// TIA Portal V20 export
// export: Created 2026-10-12T15:46:51.9760666Z, ExportSetting WithDefaults, DisplayName Totally Integrated Automation Portal, DisplayVersion V20, DisplayName TIA Portal Openness, DisplayVersion V20, DisplayName TIA Portal Teamcenter Gateway, DisplayVersion V20, DisplayName TIA Portal Version Control Interface, DisplayVersion V20, DisplayName SINAMICS Startdrive Advanced, DisplayVersion V20 SP1 Update 2, DisplayName SINAMICS Startdrive G110M, G120, G120C, G120D, G120P, G115D, DisplayVersion V20 SP1 Update 2, DisplayName SINAMICS Startdrive G130, G150, S120, S150, SINAMICS MV, G220, S200, S210, DisplayVersion V20 SP1 Update 2, DisplayName STEP 7 Professional, DisplayVersion V20, DisplayName STEP 7 Safety, DisplayVersion V20, DisplayName WinCC Basic/Comfort/Advanced, DisplayVersion V20, DisplayName WinCC Professional, DisplayVersion V20, DisplayName WinCC Unified, DisplayVersion V20
DATA_BLOCK "GDB_AccessPersistTest"   // DB15
{ S7_Optimized_Access := 'TRUE' }
VERSION : 0.1
// stored: AutoNumber true, DBAccessibleFromOPCUA true, DBAccessibleFromWebserver true, IsOnlyStoredInLoadMemory false, IsRetainMemResEnabled false, IsWriteProtectedInAS false, MemoryReserve 100
   VAR
      Operation : Int;
      Value : DInt;
      Gate : Int;
      RotateOnLogin : Bool;
      Root : String[32];
      Applied { ExternalWritable := 'False'} : Bool;
      UsersReady { ExternalWritable := 'False'} : Bool;
      UsersLost { ExternalWritable := 'False'} : Bool;
      UserGeneration { ExternalWritable := 'False'} : UDInt;
      CrcWitness { ExternalWritable := 'False'} : DWord;
      Record { ExternalAccessible := 'False'; ExternalVisible := 'False'; ExternalWritable := 'False'; S7_SetPoint := 'True'} : "ST_UserRecord";
      PolicySlot { ExternalAccessible := 'False'; ExternalVisible := 'False'; ExternalWritable := 'False'} : Int;
   END_VAR
   VAR RETAIN
      ProvisionCount { ExternalWritable := 'False'} : UDInt;
      StartupCount { ExternalWritable := 'False'} : UDInt;
   END_VAR
BEGIN
END_DATA_BLOCK
